(* IEC 61131-3 sources: nautilus/website/lessons/b1-blink/variants/bad-blinks-once, 1 file *)

(* ---- program.st ---- *)
PROGRAM Blink
VAR n : INT; flips : INT; END_VAR
n := n + 1;
IF n >= 5 AND flips < 2 THEN
    Lamp := NOT Lamp;
    flips := flips + 1;
    n := 0;
END_IF;
END_PROGRAM
